(* IEC 61131-3 sources: ControlsBenchMUSE/codesys/library/examples/mappings/tank-loop, 10 files *)

(* ---- ST_TANK_Inputs.st ---- *)
TYPE ST_TANK_Inputs :
STRUCT
    // Generated by codesys/library/scripts/cb-map.mjs 0.1.0 from mappings/tank-loop.map.json; do not edit.
    // Raw inputs in native types; the session image carries them losslessly.
    LT101_Raw : INT; // Numeric.Signed[0], 16-bit
    TT102_Raw : INT; // Numeric.Signed[1], 16-bit
    PT103_Raw : UINT; // Numeric.Unsigned[0], 12-bit
    LSH104 : BOOL; // Digital[0]
    P105_RunFB : BOOL; // Digital[1]
    FQ106_Count : UDINT; // Numeric.Unsigned[1], 32-bit
    AT107_Value : REAL; // Numeric.RealValue[0]
END_STRUCT
END_TYPE

(* ---- ST_TANK_Outputs.st ---- *)
TYPE ST_TANK_Outputs :
STRUCT
    // Generated by codesys/library/scripts/cb-map.mjs 0.1.0 from mappings/tank-loop.map.json; do not edit.
    // Application output commands in native types.
    P105_RunCmd : BOOL; // Digital[0]
    XV108_OpenCmd : BOOL; // Digital[1]
    TY102_Out : INT; // Numeric.Signed[0], 16-bit
    FCV109_Out : REAL; // Numeric.RealValue[0]
END_STRUCT
END_TYPE

(* ---- ST_TANK_Taps.st ---- *)
TYPE ST_TANK_Taps :
STRUCT
    // Generated by codesys/library/scripts/cb-map.mjs 0.1.0 from mappings/tank-loop.map.json; do not edit.
    // Read-only observation taps of internal signals.
    TIC102_SP : REAL; // Numeric.RealValue[0]
    TIC102_PV : REAL; // Numeric.RealValue[1]
    TIC102_CV : REAL; // Numeric.RealValue[2]
    TIC102_Mode : INT; // Numeric.Signed[0], 16-bit
END_STRUCT
END_TYPE

(* ---- GVL_TANK_Map.st ---- *)
{attribute 'qualified_only'}
VAR_GLOBAL CONSTANT
    // Generated by codesys/library/scripts/cb-map.mjs 0.1.0 from mappings/tank-loop.map.json; do not edit.
    // Wire identities of this machine map.
    MAP_ID : STRING(32) := 'tank-loop';
    SCHEMA_ID : UDINT := 16#908F6F3C; // raw input/output channel layout
    TAP_SCHEMA_ID : UDINT := 16#A7F251A8; // observation tap list; 0 when none
    DEFAULT_DOMAIN_ID : UDINT := 2;
    TIMEOUT_US : ULINT := 750000;
END_VAR

(* ---- MAP_TANK_Config.st ---- *)
FUNCTION MAP_TANK_Config : CB.ST_CB_Config
VAR_INPUT
    DomainId : UDINT; // one value per authority domain in the application
END_VAR
VAR
    c : CB.ST_CB_Config;
END_VAR
// Generated by codesys/library/scripts/cb-map.mjs 0.1.0 from mappings/tank-loop.map.json; do not edit.
// Session configuration for this map.
c.DomainId := DomainId;
c.SchemaId := GVL_TANK_Map.SCHEMA_ID;
c.TimeoutUs := GVL_TANK_Map.TIMEOUT_US;
c.DigitalCount := 2;
c.SignedCount := 2;
c.UnsignedCount := 2;
c.RealCount := 1;
c.SignedBits[0] := 16; // LT101_Raw
c.SignedBits[1] := 16; // TT102_Raw
c.UnsignedBits[0] := 12; // PT103_Raw
c.UnsignedBits[1] := 32; // FQ106_Count
c.RealNonFiniteAllowed[0] := TRUE; // AT107_Value
MAP_TANK_Config := c;
END_FUNCTION

(* ---- MAP_TANK_PackInputs.st ---- *)
FUNCTION MAP_TANK_PackInputs : CB.ST_CB_Image
VAR_INPUT
    Source : ST_TANK_Inputs;
END_VAR
VAR
    image : CB.ST_CB_Image;
END_VAR
// Generated by codesys/library/scripts/cb-map.mjs 0.1.0 from mappings/tank-loop.map.json; do not edit.
// Raw acquisition into the session hardware image.
image.Numeric.Signed[0] := INT_TO_DINT(Source.LT101_Raw);
image.Numeric.Signed[1] := INT_TO_DINT(Source.TT102_Raw);
image.Numeric.Unsigned[0] := UINT_TO_UDINT(Source.PT103_Raw);
image.Digital[0] := Source.LSH104;
image.Digital[1] := Source.P105_RunFB;
image.Numeric.Unsigned[1] := Source.FQ106_Count;
image.Numeric.RealValue[0] := Source.AT107_Value;
MAP_TANK_PackInputs := image;
END_FUNCTION

(* ---- MAP_TANK_PackOutputs.st ---- *)
FUNCTION MAP_TANK_PackOutputs : CB.ST_CB_Image
VAR_INPUT
    Source : ST_TANK_Outputs;
END_VAR
VAR
    image : CB.ST_CB_Image;
END_VAR
// Generated by codesys/library/scripts/cb-map.mjs 0.1.0 from mappings/tank-loop.map.json; do not edit.
// Authentic commands into an output image for the DO/AO taps.
image.Digital[0] := Source.P105_RunCmd;
image.Digital[1] := Source.XV108_OpenCmd;
image.Numeric.Signed[0] := INT_TO_DINT(Source.TY102_Out);
image.Numeric.RealValue[0] := Source.FCV109_Out;
MAP_TANK_PackOutputs := image;
END_FUNCTION

(* ---- MAP_TANK_PackTaps.st ---- *)
FUNCTION MAP_TANK_PackTaps : CB.ST_CB_Image
VAR_INPUT
    Source : ST_TANK_Taps;
END_VAR
VAR
    image : CB.ST_CB_Image;
END_VAR
// Generated by codesys/library/scripts/cb-map.mjs 0.1.0 from mappings/tank-loop.map.json; do not edit.
// Observation taps into the frame tap image; no write path exists.
image.Numeric.RealValue[0] := Source.TIC102_SP;
image.Numeric.RealValue[1] := Source.TIC102_PV;
image.Numeric.RealValue[2] := Source.TIC102_CV;
image.Numeric.Signed[0] := INT_TO_DINT(Source.TIC102_Mode);
MAP_TANK_PackTaps := image;
END_FUNCTION

(* ---- MAP_TANK_UnpackInputs.st ---- *)
FUNCTION MAP_TANK_UnpackInputs : ST_TANK_Inputs
VAR_INPUT
    Image : CB.ST_CB_Image;
END_VAR
VAR
    values : ST_TANK_Inputs;
END_VAR
// Generated by codesys/library/scripts/cb-map.mjs 0.1.0 from mappings/tank-loop.map.json; do not edit.
// Selected image back to native types; the session has enforced each width.
values.LT101_Raw := DINT_TO_INT(Image.Numeric.Signed[0]);
values.TT102_Raw := DINT_TO_INT(Image.Numeric.Signed[1]);
values.PT103_Raw := UDINT_TO_UINT(Image.Numeric.Unsigned[0]);
values.LSH104 := Image.Digital[0];
values.P105_RunFB := Image.Digital[1];
values.FQ106_Count := Image.Numeric.Unsigned[1];
values.AT107_Value := Image.Numeric.RealValue[0];
MAP_TANK_UnpackInputs := values;
END_FUNCTION

(* ---- MAP_TANK_UnpackOutputs.st ---- *)
FUNCTION MAP_TANK_UnpackOutputs : ST_TANK_Outputs
VAR_INPUT
    Image : CB.ST_CB_Image;
END_VAR
VAR
    values : ST_TANK_Outputs;
END_VAR
// Generated by codesys/library/scripts/cb-map.mjs 0.1.0 from mappings/tank-loop.map.json; do not edit.
// Physical sink values; configured SuppressedValues must fit each native type.
values.P105_RunCmd := Image.Digital[0];
values.XV108_OpenCmd := Image.Digital[1];
values.TY102_Out := DINT_TO_INT(Image.Numeric.Signed[0]);
values.FCV109_Out := Image.Numeric.RealValue[0];
MAP_TANK_UnpackOutputs := values;
END_FUNCTION
